# EPICS substitutions: db/Beckhoff_1XXX/ecmcEK1101.substitutions
file "ecmc_coupler-ID.template"
{
  pattern {}
          {}
}
